Fanuc KAREL source: KT00593.KL

PROGRAM KT00593
%NOLOCKGROUP
VAR
  I1: INTEGER
  I2: INTEGER
  OUT: STRING[80]
BEGIN
  I1 = 2
  I2 = 3
  I1 = 2
  I2 = 3
  OUT = I1 + I2
END KT00593
